// TIA Portal V20 export
// export: Created 2026-10-19T18:45:54.0218764Z, ExportSetting None, DisplayName Totally Integrated Automation Portal, DisplayVersion V20 Update 6, DisplayName TIA Portal Openness, DisplayVersion V20 Update 6, DisplayName TIA Portal Version Control Interface, DisplayVersion V20 Update 6, DisplayName SINAMICS Startdrive Advanced, DisplayVersion V20 SP1, DisplayName SINAMICS Startdrive G130, G150, S120, S150, SINAMICS MV, G220, S200, S210, DisplayVersion V20 SP1, DisplayName SINAMICS Startdrive G110M, G120, G120C, G120D, G120P, G115D, DisplayVersion V20 SP1, DisplayName STEP 7 Professional, DisplayVersion V20 Update 6, DisplayName STEP 7 Safety, DisplayVersion V20 Update 2, DisplayName WinCC Basic/Comfort/Advanced, DisplayVersion V20 Update 6, DisplayName WinCC Unified, DisplayVersion V20 Update 6
VAR_GLOBAL   // PLC tag table "IO_Charger Panel_L6"
   "CHARGER L6 - Output Current" AT %ID872 : Real;   // Actual Output Current
   "CHARGER L6 - Confirm Voltage & Current Setting" AT %Q442.2 : Bool;   // Confirmation Command
   "CHARGER L6 - Output Voltage" AT %ID868 : Real;   // Actual Output Voltage
   "CHARGER L6 - Set Current Feedback" AT %ID880 : Real;   // Set Current Value
   "CHARGER L6 - Stop Charging" AT %Q442.1 : Bool;   // Stop Charging Command
   "CHARGER L6 - Set Voltage Feedback" AT %ID876 : Real;   // Set Voltage Value
   "CHARGER L6 - Charging Start" AT %I884.0 : Bool;   // Charging Running Status
   "CHARGER L6 - Start Charging" AT %Q442.0 : Bool;   // Start Charging Command
   "CHARGER L6 - Set Current Output" AT %QD438 : Real;   // Issue Target Current
   "CHARGER L6 - Set Voltage Output" AT %QD434 : Real;   // Issue Target Voltage
END_VAR
